Fanuc KAREL source: kt00735.KL

-- PROVISIONAL review KL for V770-1; original PC SHA256 67c81b72875245aab60e19edbf03033e9bde84d2857074a7af2aad4de7823719
-- Incomplete behavior may be omitted. Consult companion uncertainty JSON. Do not deploy.
PROGRAM KT00735
%NOLOCKGROUP
VAR
  OUT : INTEGER
-- UNRESOLVED_DECL ARG type=002012
BEGIN
  -- UNRESOLVED_PC offsets 5-18; opcodes 22,1D,23
  -- UNRESOLVED_PC offsets 23-27; opcodes 7F
END KT00735
